(* IEC 61131-3 sources: teller/JD_Teller_LC2_V11/Network/JamDetection_Trombone, 1 file *)

(* ---- ONE_JamDetection_Trombone_Table.st ---- *)
#define OBJECTS_CONFIG

FUNCTION GLOBAL TAB ONE_JamDetection_Trombone
-1$UINT, 0$UINT,
0$UINT, 0$UINT,

9$UDINT,
TO_UDINT(800276940), "_AlarmX0Para", 0$UINT, 4$UINT, 0$UINT,
TO_UDINT(1746090780), "_AlarmX3Para", 0$UINT, 2$UINT, 1$UINT,
TO_UDINT(3293687312), "Call_JAM_Window", 1$UINT, 0$UINT, 1$UINT,
TO_UDINT(2466162658), "JAMDETECT_Teller", 1$UINT, 0$UINT, 1$UINT,
TO_UDINT(826277511), "Jamdetection_TeachIn_Teller", 1$UINT, 1$UINT, 1$UINT,
TO_UDINT(2225119864), "MerkerEx", 1$UINT, 18$UINT, 0$UINT,
TO_UDINT(933570811), "RAMex", 1$UINT, 16$UINT, 1$UINT,
TO_UDINT(1060418456), "Signal_Splitter_BG_Teller", 1$UINT, 0$UINT, 1$UINT,
TO_UDINT(1383955435), "Visu_Jam", 0$UINT, 0$UINT, 3$UINT,

_NO_ATTR, TO_UDINT(604600958), "JAMDETECT_ALARM",

_NO_ATTR, TO_UDINT(2662313597), "CALL_JAM_WINDOW1",

_NO_ATTR, TO_UDINT(1648271141), "JAMDETECT1",

_NO_ATTR, TO_UDINT(3822706166), "S11_JAMDETECTION_TEACHIN_01",

_NO_ATTR, TO_UDINT(2288677303), "S11_RAM_JAMDETECTION_TEACHIN_01",

_NO_ATTR, TO_UDINT(550170101), "VISU_TEACHIN_JAMDETECT",

_NO_ATTR, TO_UDINT(2438206062), "S11_VISUJAMDETECT_01",
_NO_ATTR, TO_UDINT(140329940), "S11_VISUJAMDETECT_02",
_NO_ATTR, TO_UDINT(2136634178), "S11_VISUJAMDETECT_03",

//Internal connections
0$UDINT,
0$UDINT,
0$UDINT,
12$UDINT,
TO_UDINT(0), "Para1", TO_UDINT(2), "Jam_ID_Section",
TO_UDINT(0), "Para2", TO_UDINT(2), "Jam_ID_Unit",
TO_UDINT(0), "Para3", TO_UDINT(2), "Jam_Count",
TO_UDINT(2), "cJamReset", TO_UDINT(3), "ResetJam",
TO_UDINT(2), "cJam_Trombone", TO_UDINT(4), "m_udLength",
TO_UDINT(2), "cJamLSE", TO_UDINT(1), "ClassSvr",
TO_UDINT(2), "Jam2Visu", TO_UDINT(0), "ClassSvr",
TO_UDINT(3), "c_JamData", TO_UDINT(4), "m_udLength",
TO_UDINT(5), "c_WriteValue01", TO_UDINT(3), "TeachIn",
TO_UDINT(6), "c_JamData", TO_UDINT(4), "m_udLength",
TO_UDINT(7), "c_JamData", TO_UDINT(4), "m_udLength",
TO_UDINT(8), "c_JamData", TO_UDINT(4), "m_udLength",

//Initialization values
0$UDINT,
10$UDINT,
TO_UDINT(0), "Config", TO_UDINT(0),//|JamDetection_Trombone.JAMDETECT_ALARM.Config;
TO_UDINT(2), "JamResetC001", TO_UDINT(0),//|JamDetection_Trombone.JAMDETECT1.JamResetC001;
TO_UDINT(2), "Jam2Visu", TO_UDINT(0),//|JamDetection_Trombone.JAMDETECT1.Jam2Visu;
TO_UDINT(3), "c_SectieType", TO_UDINT(11),//|JamDetection_Trombone.S11_Jamdetection_TeachIn_01.c_SectieType;
TO_UDINT(3), "cJamDetect2HW", TO_UDINT(0),//|JamDetection_Trombone.S11_Jamdetection_TeachIn_01.cJamDetect2HW;
TO_UDINT(3), "cJamReset", TO_UDINT(0),//|JamDetection_Trombone.S11_Jamdetection_TeachIn_01.cJamReset;
TO_UDINT(4), "ThreadSafe", TO_UDINT(0),//|JamDetection_Trombone.S11_RAM_Jamdetection_TeachIn_01.ThreadSafe;
TO_UDINT(6), "c_SensorNr", TO_UDINT(1),//|JamDetection_Trombone.S11_VisuJamdetect_01.c_SensorNr;
TO_UDINT(7), "c_SensorNr", TO_UDINT(2),//|JamDetection_Trombone.S11_VisuJamdetect_02.c_SensorNr;
TO_UDINT(8), "c_SensorNr", TO_UDINT(3),//|JamDetection_Trombone.S11_VisuJamdetect_03.c_SensorNr;

//Symbolic initialization values
0$UDINT,
0$UDINT,

//Initialization of string values
0$UDINT,
0$UDINT,

//Configuration of tasks (RealTime, Cyclic, Background)
0$UDINT,
1$UDINT,
TO_UDINT(3), (1)$UDINT, 4194305$DINT, 	//S11_JAMDETECTION_TEACHIN_01

0$UDINT,
2$UDINT,
TO_UDINT(2), (100)$UDINT, 4194305$DINT, 	//JAMDETECT1
TO_UDINT(3), (50)$UDINT, 4194305$DINT, 	//S11_JAMDETECTION_TEACHIN_01

0$UDINT,
4$UDINT,
TO_UDINT(5), (100)$UDINT, 4194305$DINT, 	//VISU_TEACHIN_JAMDETECT
TO_UDINT(6), (100)$UDINT, 4194305$DINT, 	//S11_VISUJAMDETECT_01
TO_UDINT(7), (100)$UDINT, 4194305$DINT, 	//S11_VISUJAMDETECT_02
TO_UDINT(8), (100)$UDINT, 4194305$DINT, 	//S11_VISUJAMDETECT_03

//External connections
0$UDINT,
7$UDINT,
TO_UDINT(2), "JamResetTanabe", C_TRY, TO_UDINT(396609901), "CIO011_IM1","Input6",
TO_UDINT(2), "JamKlok", C_TRY, TO_UDINT(2236149643), "SerSend1","Jamdetect",
TO_UDINT(3), "iEncoder", C_TRY, TO_UDINT(396609901), "CIO011_IM1","Encoder",
TO_UDINT(3), "cJamDetect2HW", C_DIR, TO_UDINT(2206833861), "JD_OR1","In2",
TO_UDINT(3), "cSensor_01", C_TRY, TO_UDINT(396609901), "CIO011_IM1","Input4",
TO_UDINT(3), "cSensor_02", C_TRY, TO_UDINT(396609901), "CIO011_IM1","Input5",
TO_UDINT(3), "cSensor_03", C_TRY, TO_UDINT(396609901), "CIO011_IM1","Input3",

//Magic internal connections
0$UDINT,
0$UDINT,

//Configuration of timeslots of tasks (RealTime, Cyclic)
#ifdef __LSLLDR_TIMESLOTS__
0$UDINT,
0$UDINT,

0$UDINT,
0$UDINT,

#endif //__LSLLDR_TIMESLOTS__

//MultiMaster connections
#ifdef __LSLLDR_MULTIMASTER__
0$UDINT,
0$UDINT,
#endif //__LSLLDR_MULTIMASTER__

END_FUNCTION
